Fanuc KAREL source: kc00038.KL

-- PROVISIONAL review KL for V1013-1; original PC SHA256 3f3a8b592a80096685babe260b5f497865eddc28cb067071a88dc6dc815abffd
-- Incomplete behavior may be omitted. Consult companion uncertainty JSON. Do not deploy.
PROGRAM KC00038
%NOLOCKGROUP
BEGIN
  -- UNRESOLVED_PC offsets 5-32; opcodes 27,22,1C,22,22,76
  -- UNRESOLVED_PC offsets 37-41; opcodes 7F
END KC00038
